(* Schneider Machine Expert - Basic project Case01, file version 2.9.0.0 *)
(* ProjectInformations: Name=New project *)

HARDWARE
  Cpu 0: TM221M16R/G
  EthernetConfiguration: NetworkName=M221, IpAllocationMode=FixedAddress, IpAddress=0.0.0.0, SubnetMask=0.0.0.0
  SerialLineConfiguration: Baud=Baud19200, Parity=ParityEven, DataBits=DataBits8, StopBits=StopBits1, PhysicalMedium=PhysicalMediumRs485, TransmissionMode=TransmissionModeModbusRtu, SlaveId=1, Addressing=SlaveAddressing
  MastTask: UsePeriodScanMode=false, PeriodScan=100
  FastTask: Period=255
  CpuBehavior: StartingMode=StartAsPreviousState, AutoSaveRamOnEeprom=true, WatchdogPeriod=250

SYMBOLS  (address, symbol, comment, settings)
  %M0       Armed
  %M1       RunRequest
  %TM0        [Preset=3, Base=OneSecond]
  %I0.0     StartPB
  %I0.1     StopHealthy
  %I0.2     EStopHealthy
  %I0.3     GuardHealthy
  %Q0.0     Motor
  %Q0.1     Horn

POU New POU
  (* SectionNumber=1 *)

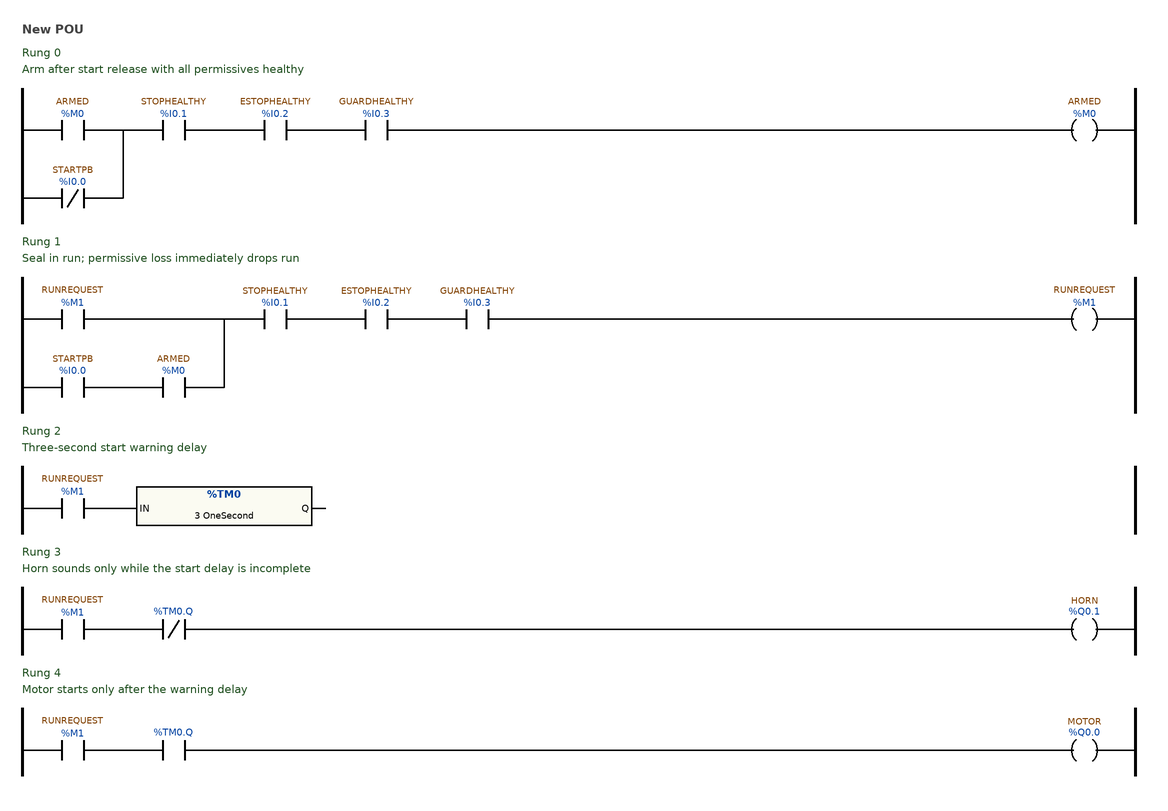

// Rung 0
// Arm after start release with all permissives healthy
  LD %M0                  (* Armed *)
  ORN %I0.0               (* StartPB *)
  AND %I0.1               (* StopHealthy *)
  AND %I0.2               (* EStopHealthy *)
  AND %I0.3               (* GuardHealthy *)
  ST %M0                  (* Armed *)
  // as ST:
  //   Armed := (Armed OR NOT StartPB) AND StopHealthy AND EStopHealthy AND GuardHealthy;

// Rung 1
// Seal in run; permissive loss immediately drops run
  LD %M1                  (* RunRequest *)
  OR( %I0.0               (* StartPB *)
  AND %M0                 (* Armed *)
  )
  AND %I0.1               (* StopHealthy *)
  AND %I0.2               (* EStopHealthy *)
  AND %I0.3               (* GuardHealthy *)
  ST %M1                  (* RunRequest *)
  // as ST:
  //   RunRequest := (RunRequest OR StartPB AND Armed) AND StopHealthy AND EStopHealthy AND GuardHealthy;

// Rung 2
// Three-second start warning delay
  BLK %TM0
  LD %M1                  (* RunRequest *)
  IN
  END_BLK
  // as ST:
  //   %TM0(IN := RunRequest);

// Rung 3
// Horn sounds only while the start delay is incomplete
  LD %M1                  (* RunRequest *)
  ANDN %TM0.Q
  ST %Q0.1                (* Horn *)
  // as ST:
  //   Horn := RunRequest AND NOT %TM0.Q;

// Rung 4
// Motor starts only after the warning delay
  LD %M1                  (* RunRequest *)
  AND %TM0.Q
  ST %Q0.0                (* Motor *)
  // as ST:
  //   Motor := RunRequest AND %TM0.Q;
